(* CODESYS project keyence_sr.library
   Company: KOSTAL GmbH & Co.KG
   Version: 1.0.0.0
   DefaultNamespace: KOSTAL.AF2024.Drivers.Scanner.Keyence_SR
   Title: KOSTAL.AF2024.Drivers.Scanner.Keyence_SR
   Placeholder: KOSTAL.AF2024.Drivers.Scanner.Keyence_SR
   Author: Frank Dümpelmann
   DocFormat: reStructuredText

Project tree, tasks and I/O mapping:
  libraries: KOSTAL.AF2024.Core.ListOf, 1.0.0.0 (KOSTAL GmbH & Co.KG); KOSTAL.AF2024.Core.Process, 1.0.0.0 (KOSTAL GmbH & Co.KG); KOSTAL.AF2024.Core.Settings, 1.0.0.0 (KOSTAL GmbH & Co.KG); KOSTAL.AF2024.Core.StringTools, 1.0.0.0 (KOSTAL GmbH & Co.KG); KOSTAL.AF2024.Drivers.Scanner.IScanner, 1.0.0.0 (KOSTAL GmbH & Co.KG); Tc2_Standard, 3.3.3.0 (Beckhoff Automation GmbH); Tc2_TcpIp, 3.3.10.0 (Beckhoff Automation GmbH)
  DUT/
    data type E_PROCESS
  EthernetIP/
    DUTs/
      data type ST_SR751_IN
      data type ST_SR751_OUT
    function block FB_Reader_EthernetIP [ST]: ClearCodes, CodeGet, Ex_Scan, NativeStringGet, NumberOfBarcodes, State, _0_ready, _1_finish, _2_analyseResponse, _2_read, _2_split, _connectControl, _FBmain, FB_init, FBmain
  Project Information/
    function F_GetCompany [ST]
    function F_GetTitle [ST]
    function F_GetVersion [ST]
  TCP_IP/
    function block FB_Reader_TcpIp [ST]: ClearCodes, CodeGet, Ex_Scan, NativeStringGet, NumberOfBarcodes, State, _devices, _FBmain, _splitString, _stepConnect, _stepFinish, _stepReady, _stepReceive, _stepSend, _timeOutOccured, Command, ETX, ExecutedSocketState, intermediateLimiter, remote_IP, remote_Port, separator, serverAmsNetId, STX, timeOut, FB_init, FBmain
    interface I_Scanner: ExecutedSocketState
  Version/
    global variables Global_Version
*)

// DUT/E_PROCESS
{attribute 'qualified_only'}
{attribute 'strict'}
TYPE E_PROCESS :
(
	idle			:= 0,
	scan	:= 1
);
END_TYPE

// EthernetIP/DUTs/ST_SR751_IN
{attribute 'pack_mode' := '1'} 
TYPE ST_SR751_IN :
	STRUCT
		Error	: BIT;
		ResultDataAvailable	: BIT;
		ResultDataStrobe	: BIT;
		noName_0_0	: BIT;
		noName_0_1	: BIT;
		noName_0_2	: BIT;
		BufferOverfolwError	: BIT;
		GeneralError	: BIT;
		Busy	: BIT;
		TRG_BUSY	: BIT;
		LOCK_BUSY	: BIT;
		MODE_BUSY	: BIT;
		ERR_BUSY	: BIT;
		noName_1_0	: BIT;
		noName_1_1	: BIT;
		noName_1_2	: BIT;
		ReadComplete	: BIT;
		PresetComplete	: BIT;
		RegisterPresetDataComplete	: BIT;
		TuneComplete	: BIT;
		noName_2_0	: BIT;
		noName_2_1	: BIT;
		noName_2_2	: BIT;
		EXT_RequestComplete	: BIT;
		ReadFailure	: BIT;
		PresetFailure	: BIT;
		RegisterPresetDataFailure	: BIT;
		TuneFailure	: BIT;
		noName_3_0	: BIT;
		noName_3_1	: BIT;
		noName_3_2	: BIT;
		EXT_RequestFailure	: BIT;
		IN_1_Status	: BIT;
		IN_2_Status	: BIT;
		noName_4_0	: BIT;
		noName_4_1	: BIT;
		OUT_1_Status	: BIT;
		OUT_2_Status	: BIT;
		OUT_3_Status	: BIT;
		noName_5	: BIT;
		Unstable	: BIT;
		MatchingLevelUnstable	: BIT;
		ISO_IEC_15415_Unstable	: BIT;
		AIM_DPM_Unstable	: BIT;
		SAE_A59132_Unstable	: BIT;
		noName_6_0	: BIT;
		noName_6_1	: BIT;
		noName_6_2	: BIT;
		noName_6_3	: BIT;
		noName_6_4	: BIT;
		noName_6_5	: BIT;
		noName_6_6	: BIT;
		noName_6_7	: BIT;
		noName_6_8	: BIT;
		noName_6_9	: BIT;
		noName_6_10	: BIT;
		noName_6_11	: BIT;
		noName_6_12	: BIT;
		noName_6_13	: BIT;
		noName_6_14	: BIT;
		noName_6_15	: BIT;
		noName_6_16	: BIT;
		noName_6_17	: BIT;
		noName_6_18	: BIT;
		MatchingLevel	: UINT;
		ISO_IEC_15415_Grade	: UINT;
		AIM_DPM_Grade	: UINT;
		noName_7	: ARRAY[0..1] OF BYTE;
		ReadResultCode	: UINT;
		PresetResultCode	: UINT;
		RegisterPresetDataResultCode	: UINT;
		TuneResultCode	: UINT;
		noName_8	: ARRAY[0..5] OF BYTE;
		EXT_RequestResultCode	: UINT;
		GeneralErrorCode	: UINT;
		noName_9	: ARRAY[0..1] OF BYTE;
		ResultDataReadyCount	: UINT;
		ResultDataUpdateCount	: UINT;
		noName_10	: ARRAY[0..1] OF BYTE;
		ResultDataSize	: UINT;
		ResultData : STRING(81);
		
		
		
		
	END_STRUCT
END_TYPE

// EthernetIP/DUTs/ST_SR751_OUT

TYPE ST_SR751_OUT :
	STRUCT
		noName0_BIT	: BIT;
		ResultDataLatch	: BIT;
		noName_1_0	: BIT;
		noName_1_1	: BIT;
		noName_1_2	: BIT;
		noName_1_3	: BIT;
		noName_1_4	: BIT;
		ErrorClear	: BIT;
		ReadRequest	: BIT;
		PresetRequest	: BIT;
		RegisterPresetDataRequest	: BIT;
		TuneRequest	: BIT;
		noName_2_0	: BIT;
		noName_2_1	: BIT;
		noName_2_2	: BIT;
		noName_2_3	: BIT;
		ReadCompleteClear	: BIT;
		PresetCompleteClear	: BIT;
		RegisterPresetDataCompleteClear	: BIT;
		TuneCompleteClear	: BIT;
		noName_3_0	: BIT;
		noName_3_1	: BIT;
		noName_3_2	: BIT;
		ExtRequestCompleteClear	: BIT;
		noName_4	: BYTE;
		BankNumber	: UINT;
		noName_5_0	: BYTE;
		noName_5_1	: BYTE;
		noName_5_2	: BYTE;
		noName_5_3	: BYTE;
		UserDataSize:	UINT;
		UserData	: ARRAY[14..77] OF BYTE;
	END_STRUCT
END_TYPE

// Version/Global_Version
{attribute 'TcGenerated'}
{attribute 'no-analysis'}
{attribute 'linkalways'}
// This function has been automatically generated from the project information.
VAR_GLOBAL CONSTANT
	{attribute 'const_non_replaced'}
	stLibVersion_KOSTAL_AF2024_Drivers_Scanner_Keyence_SR : ST_LibVersion := (iMajor := 1, iMinor := 0, iBuild := 0, iRevision := 0, nFlags := 0, sVersion := '1.0.0.0');
END_VAR

// EthernetIP/FB_Reader_EthernetIP
(*
From EDS Specification Keyence_1003_0101.eds from 22.11.2012 12:56
===================================================================
*)

FUNCTION_BLOCK FB_Reader_EthernetIP IMPLEMENTS KOSTAL_AF2024_Drivers_Scanner_IScanner.I_Scanner



VAR
	ECatState	AT %I*	: UINT;	//link to EtherCat State from {Device x (ECAT EIP Scanner (EL6652))}.Inputs.State
	SR_750_Series_State	AT %I*	: UINT;	//link to {SR-750 Series}.Inputs.State

	SR751_IN	AT %I*	: ARRAY[2..173] OF BYTE; //link with Continious mode ATTENTION be sure, that the Array-Nodes are collapsed
	SR751_OUT	AT %Q*	: ARRAY[2..77] OF BYTE; //link with Continious mode ATTENTION be sure, that the Array-Nodes are collapsed
	
	_pIN		: POINTER TO ST_SR751_IN;
	_pOUT	: POINTER TO ST_SR751_OUT;

	//
	_step		: KOSTAL_AF2024_Core_Process.FB_processStep;
	_THIS_CALLED			: E_PROCESS;
	_THIS_IN_PROCESS		: E_PROCESS;
	_state 	: KOSTAL_AF2024_Core_Process.T_plcState;

	//
	_split	: Kostal_AF2024_Core_StringTools.FB_Split_UTF8;
	_barcodes	: KOSTAL_AF2024_Core_ListOf.FB_ListOfString_UTF8;
	
	_nativeResult	: KOSTAL_AF2024_Core_Settings.T_MaxString_UTF8;
	

	
END_VAR

VAR CONSTANT
	_DELIMITER	: STRING(1):= '$1D';
	_STX	: STRING(1):= '$02';
	_ETX	: STRING(1):= '$03';
	_CR	: STRING(1):= '$0D';
	_LF	: STRING(1):= '$0A';
END_VAR

METHOD ClearCodes

_barcodes.clear();
_nativeResult := '';
END_METHOD

METHOD CodeGet : STRING(255)
VAR_INPUT
	number	: UINT;
END_VAR
CodeGet:= _barcodes.line_GET(number);
END_METHOD

METHOD Ex_Scan : BOOL
IF _THIS_CALLED <> E_PROCESS.idle THEN //Another process is running: don't start this process!
	Ex_Scan:= FALSE;	
	RETURN; 
END_IF


_THIS_CALLED := E_PROCESS.scan;

_FBmain();	//Call sequence via _FBmain

Ex_Scan := _THIS_CALLED = _THIS_IN_PROCESS;	//Return true when process was started
END_METHOD

METHOD NativeStringGet : STRING(255)
NativeStringGet:= _nativeResult;
END_METHOD

PROPERTY PUBLIC NumberOfBarcodes : UDINT
GET
NumberOfBarcodes:= _barcodes.NumberOfLines;
END_GET
END_PROPERTY

PROPERTY State : KOSTAL_AF2024_Core_Process.I_T_plcState
GET

State := _state;
END_GET
END_PROPERTY

METHOD PROTECTED _0_ready
VAR_INPUT
END_VAR


IF _pOUT^.ReadRequest THEN _pOUT^.ReadRequest:= FALSE;	END_IF
_pOUT^.ReadCompleteClear:= _pIN^.ReadComplete OR _pIN^.ReadFailure;
 
_state.clear();

IF _pIN^.ReadComplete OR _pIN^.ReadFailure THEN
	_state.busy := TRUE;
	_state.description:= "wait until Scanner is not longer busy";
ELSE
	_step.INC();
END_IF
END_METHOD

METHOD PROTECTED _1_finish
VAR_INPUT
END_VAR

_state.clear();

_state.finish := TRUE;
_state.pass:= TRUE;

//IF NOT _startProcess THEN	_step.set(0);	END_IF
END_METHOD

METHOD PROTECTED _2_analyseResponse
VAR_INPUT
END_VAR

_pOUT^.ReadRequest:= FALSE;
 
_state.clear();
_state.busy := TRUE;

IF NOT _pIN^.ReadFailure THEN

	_step.INC();


ELSE
	
	
	_state.finish := TRUE;
	_state.fail:= TRUE;
	_state.description:= STRING_TO_WSTRING(_pIN^.ResultData);

END_IF
END_METHOD

METHOD PROTECTED _2_read
VAR_INPUT
END_VAR


_pOUT^.ReadRequest:= TRUE;
 
_state.clear();
_state.busy := TRUE;

IF NOT _pIN^.ReadComplete THEN

	_state.description:= "wait until Scanner is finish";
	
ELSE
	
	_nativeResult:= _pIN^.ResultData;
	_step.INC();
	
END_IF
END_METHOD

METHOD PROTECTED _2_split
VAR_INPUT
END_VAR

VAR
	_i: UDINT;
	_replace: STRING(255);
END_VAR


_split.clear();
_split.Delimiter:= _DELIMITER;
_split.split(_nativeResult);
_barcodes.clear();

FOR _i:= 1 TO _split.Results.NumberOfLines DO

	_replace:= _split.Results.line_GET(_i);

	IF _replace <> '' THEN
		_replace:= Kostal_AF2024_Core_StringTools.F_Replace_UTF8(source:= _replace,toReplace:= _STX, replaceWith:= '', numberOfReplaces:= -1);
		_replace:= Kostal_AF2024_Core_StringTools.F_Replace_UTF8(source:= _replace,toReplace:= _ETX, replaceWith:= '', numberOfReplaces:= -1);
		_replace:= Kostal_AF2024_Core_StringTools.F_Replace_UTF8(source:= _replace,toReplace:= _CR, replaceWith:= '', numberOfReplaces:= -1);
		_replace:= Kostal_AF2024_Core_StringTools.F_Replace_UTF8(source:= _replace,toReplace:= _LF, replaceWith:= '', numberOfReplaces:= -1);
		_barcodes.addLine(_replace);
		
	END_IF

END_FOR

_step.INC();
END_METHOD

METHOD PROTECTED _connectControl : BOOL
VAR_INPUT
END_VAR

 
IF ECatState <> 0  THEN

	_connectControl:= FALSE;

	_state.clear();
	_state.fail:= TRUE;
	_state.description:= Tc2_Standard.WCONCAT(UINT_TO_WSTRING(ECatState), ";Error from EtherCAT (EIP-Scanner)");


	_step.init();

ELSIF SR_750_Series_State <> 0 THEN

	_connectControl:= FALSE;

	_state.clear();
	_state.fail:= TRUE;
	_state.description:= Tc2_Standard.WCONCAT(UINT_TO_WSTRING(SR_750_Series_State), ";Error from Ethernet IP Connection");

	_step.init();

ELSE
	
	_connectControl:= TRUE;

END_IF
END_METHOD

METHOD PROTECTED _FBmain
VAR_INPUT
END_VAR

_pIN:= ADR(SR751_IN[2]);
_pOUT:= ADR(SR751_OUT[2]);


IF NOT _connectControl() THEN RETURN;	END_IF

IF _THIS_CALLED <> _THIS_IN_PROCESS THEN
	_step.init();
END_IF

_THIS_IN_PROCESS:= _THIS_CALLED;

IF _THIS_CALLED = E_PROCESS.scan THEN

	_step.Header();
	
	CASE _step.actual OF
		
		0:	_0_ready();
		1:	_2_read();
		2:	_2_analyseResponse();
		3:	_2_split();
		4:	_1_finish();
		
	ELSE
		
		_state.clear();
		_state.fail:= TRUE;
		_state.description:= Tc2_Standard.WCONCAT(INT_TO_WSTRING(_step.actual), ". Step does not exist");
		
	END_CASE

ELSE
	_state.clear();
	_state.ready := TRUE;
END_IF
END_METHOD

METHOD FB_init : BOOL
VAR_INPUT
	bInitRetains : BOOL; // if TRUE, the retain variables are initialized (warm start / cold start)
	bInCopyCode : BOOL;  // if TRUE, the instance afterwards gets moved into the copy code (online change)
END_VAR

_pIN:= ADR(SR751_IN[2]);
_pOUT:= ADR(SR751_OUT[2]);
END_METHOD

METHOD PUBLIC FBmain
VAR_INPUT
END_VAR
IF _THIS_CALLED = E_PROCESS.idle THEN
	_FBmain();
END_IF

_THIS_CALLED:= E_PROCESS.idle;
END_METHOD

END_FUNCTION_BLOCK

// TCP_IP/I_Scanner
INTERFACE I_Scanner EXTENDS KOSTAL_AF2024_Drivers_Scanner_IScanner.I_Scanner

(*
Description
===========
| State of the TCP/IP connection
*)
PROPERTY PUBLIC ExecutedSocketState : E_SocketConnectionState
GET
END_GET
END_PROPERTY

END_INTERFACE

// Project Information/F_GetCompany
// This function has been automatically generated from the project information.
{attribute 'signature_flag' := '1073741824'}
{attribute 'TcGenerated'}
{attribute 'no-analysis'}
FUNCTION F_GetCompany : WSTRING
VAR_INPUT
	
END_VAR

F_GetCompany := "KOSTAL GmbH & Co.KG";

END_FUNCTION

// Project Information/F_GetTitle
// This function has been automatically generated from the project information.
{attribute 'signature_flag' := '1073741824'}
{attribute 'TcGenerated'}
{attribute 'no-analysis'}
FUNCTION F_GetTitle : WSTRING
VAR_INPUT
	
END_VAR

F_GetTitle := "KOSTAL.AF2024.Drivers.Scanner.Keyence_SR";

END_FUNCTION

// Project Information/F_GetVersion
// This function has been automatically generated from the project information.
{attribute 'signature_flag' := '1073741824'}
{attribute 'TcGenerated'}
{attribute 'no-analysis'}
FUNCTION F_GetVersion : ST_LibVersion
VAR_INPUT
	
END_VAR

F_GetVersion.iMajor := 1;
F_GetVersion.iMinor := 0;
F_GetVersion.iBuild := 0;
F_GetVersion.iRevision := 0;
F_GetVersion.sVersion := '1.0.0.0';
F_GetVersion.nFlags := 0;

END_FUNCTION

// TCP_IP/FB_Reader_TcpIp
{info 'The Beckhoff Library >TF6310-TCP-IP.exe< is needed'}
(*

:Author: Frank Dümpelmann <f.duempelmann@kostal.com>, Martin Hundt <m.hundt@kostal.com>
:Date: 2019-01-07

Function
========
| Extension of FB_Reader to connect to a barcode reader via TCP/IP
| Tested with Keyence SR 750 

Usage notes
===============
| Asyncronous function block: FBmain() method must be called cyclicly
| The Beckhoff Library >TF6310-TCP-IP.exe< is needed
| 	_mode_SR750	:	BOOL;	// use this mode with KEYENCE SR 750, because the command Acknowlede is not possible to disable.

Methods and Properties
======================
| See bottom of this document for a detailed description of each method or property
| Methods starting with an underline(_) are internally used and can be ignored by the user

| Usage sample: ..\Device\Scanner\scannerBestPractice
| Usage Keyence Template ..\Device\Scanner\Keyence_SR\Keyence SR-750.ptc .. \Keyence SR-1000.ptc

*)
FUNCTION_BLOCK PUBLIC FB_Reader_TcpIp  IMPLEMENTS I_Scanner
VAR_INPUT
END_VAR
VAR_OUTPUT
END_VAR

VAR
	

	_step			: KOSTAL_AF2024_Core_Process.FB_processStep;	
	_THIS_CALLED			: E_PROCESS;
	_THIS_IN_PROCESS		: E_PROCESS;
	            	
	_state 			: KOSTAL_AF2024_Core_Process.T_plcState;
	            	
	_Command		: STRING;	//STRING to define in FB_init()
	_STX			: STRING;	//STRING to define in FB_init()
	_ETX			: STRING;	//STRING to define in FB_init()
	_timeOut		: TIME	;	//TIME to define in FB_init()
	
	_receivedString	: KOSTAL_AF2024_Core_Settings.T_MaxString_UTF8;
	_split			: Kostal_AF2024_Core_StringTools.FB_Split_UTF8;
	_barcodes		: KOSTAL_AF2024_Core_ListOf.FB_ListOfString_UTF8;

	_serverAmsNetId	: STRING:= '';	//STRING:= '' - default on local system
	_remote_IP			: STRING;	//STRING
	_remote_Port		: UDINT:= 9004;	//UDINT

	_socket				: Tc2_TcpIp.FB_ClientServerConnection;	//Tc2_TcpIp.FB_ClientServerConnection
	_executedSocketState	:	E_SocketConnectionState;
	
	_send			: Tc2_TcpIp.FB_SocketSend;	//Tc2_TcpIp.FB_SocketSend
	_receive	: Tc2_TcpIp.FB_SocketReceive;	//Tc2_TcpIp.FB_SocketReceive
	_receiveComponent	: STRING(255);	//STRING(255)
	_receiveAck	: STRING(255);	//STRING(255)

	_timeOutTimer	: TON;	//TON

	_intermediateLimiter	: STRING(1):= '$1D';
	_separator						: STRING(1):= '$1E';
	
	_subStep	: KOSTAL_AF2024_Core_Process.FB_processStep;
	_concat	: Kostal_AF2024_Core_StringTools.FB_Concat;
	
	
	

END_VAR

METHOD ClearCodes

_barcodes.clear();
_receivedString := '';
END_METHOD

(*
Description
===========
| get barcode element (number)
*)
METHOD CodeGet : KOSTAL_AF2024_Core_Settings.T_MaxString_UTF8
VAR_INPUT
	number	: UINT;
END_VAR
IF (number = 0) OR (number > _barcodes.numberOfLines) THEN
	CodeGet:= '';
ELSE
	CodeGet:= _barcodes.line_GET(number);
END_IF
END_METHOD

METHOD Ex_Scan : BOOL
IF _THIS_CALLED <> E_PROCESS.idle THEN //Another process is running: don't start this process!
	Ex_Scan:= FALSE;	
	RETURN; 
END_IF


_THIS_CALLED := E_PROCESS.scan;

_FBmain();	//Call sequence via _FBmain

Ex_Scan := _THIS_CALLED = _THIS_IN_PROCESS;	//Return true when process was started
END_METHOD

METHOD NativeStringGet : STRING(255)
NativeStringGet:= _receivedString;
END_METHOD

PROPERTY NumberOfBarcodes : UDINT
GET
NumberOfBarcodes:= _barcodes.NumberOfLines;
END_GET
END_PROPERTY

(*
Description
===========
| Status of the block
*)
PROPERTY PUBLIC State : KOSTAL_AF2024_Core_Process.I_T_plcState
GET


State := _state;
END_GET
END_PROPERTY

METHOD PROTECTED _devices
VAR_INPUT
END_VAR


_timeOutTimer(IN:= , PT:= _timeOut, Q=> , ET=> );

_socket
	(
		sSrvNetID	:= _serverAmsNetId, 
		nMode			:= Tc2_TcpIp.CONNECT_MODE_ENABLEDBG, 

		sRemoteHost	:= _remote_IP, 
		nRemotePort	:= _remote_Port, 

		bEnable			:= , 
		tReconnect	:= _timeOut, 

		bBusy		=> , 
		bError	=> , 
		nErrId	=> , 
		hSocket	=> , 
		eState	=> 
	);
	
IF _socket.bEnable THEN	_executedSocketState:= _socket.eState;	END_IF
	
_send
	(
		sSrvNetId	:= _serverAmsNetId, 
		hSocket		:= _socket.hSocket, 
		cbLen			:= INT_TO_UDINT(Tc2_Standard.LEN(_Command)), 
		pSrc			:= ADR(_Command), 
		bExecute	:= , 
		tTimeout	:= _timeOut, 

		bBusy			=> , 
		bError		=> , 
		nErrId		=> 
	);
	
	
	_receive
	(
		sSrvNetId	:= _serverAmsNetId, 
		hSocket		:= _socket.hSocket, 

		cbLen:= SIZEOF(_receiveComponent) - 1, 
		pDest:= ADR(_receiveComponent), 

		bExecute:= , 
		tTimeout:= _timeOut, 

		bBusy			=> , 
		bError		=> , 
		nErrId		=> , 
		nRecBytes	=> 
	);
END_METHOD

(*
Decription
==========
| To be called cyclicly, e.g. in DeviceDefine
*)
METHOD PROTECTED _FBmain
VAR_INPUT
END_VAR
IF _THIS_CALLED <> _THIS_IN_PROCESS THEN
	_step.init();
END_IF

_THIS_IN_PROCESS:= _THIS_CALLED;

IF _THIS_CALLED = E_PROCESS.scan THEN
	_step.Header();
	
	CASE _step.actual OF
	
		0:	_stepReady();
		1:	_stepConnect();
		2:	_stepSend();
		3:	_stepReceive();
		4:	_stepFinish();
	
	ELSE
		
		_state.clear();
		_state.description:= Tc2_Standard.WCONCAT("Step does not exist", INT_TO_WSTRING(_step.actual));
		_state.fail		:= TRUE;
		_state.finish	:= TRUE;
	
	END_CASE

ELSE
	_step.init();
	_state.clear();
	_state.ready := TRUE;
END_IF
_devices();
END_METHOD

(*
| split received string depends of STX ETX
*)
METHOD PROTECTED _splitString  : BOOL

VAR
	_i: UDINT;
	_element: STRING(255);
	_stxPos: INT;
	_code: STRING(255);
END_VAR


_barcodes.clear();

IF _receivedString = '' THEN
	
	;	// no splitting possible

	
// if EXT is defined
// ============================================================================
ELSIF _ETX <> '' THEN

	_split.clear();
	_split.Delimiter:= _ETX;
	_split.Split(_receivedString);

	// if additional STX is defined then select
	IF _STX <> '' THEN

		FOR _i:= 1 TO _split.Results.NumberOfLines DO
			
			_element:= _split.Results.line_GET(_i);
			_stxPos:= Tc2_Standard.FIND(STR1:= _element, STR2:= _STX);

			IF _stxPos > 0 THEN
				_barcodes.addLine(newLine:= Tc2_Standard.RIGHT(STR:= _element, SIZE:= Tc2_Standard.LEN( STR:= _element) - _stxPos ));
			END_IF
		END_FOR
	
	// no STX defined
	ELSE

		FOR _i:= 1 TO _split.Results.NumberOfLines DO
			_barcodes.addLine(_split.Results.line_GET(_i));
		END_FOR
	
	END_IF

	
// if only STX is defined
// ============================================================================
ELSIF _STX <> '' THEN
	
	_split.clear();
	_split.Delimiter:= _STX;
	_split.Split(_receivedString);

	FOR _i:= 1 TO _split.Results.NumberOfLines DO
		_barcodes.addLine(_split.Results.line_GET( _i));
	END_FOR

// neither STX or ETX is defined then no splitting possible
// ============================================================================
ELSE

	_barcodes.addLine(newLine:= _receivedString);

END_IF

_splitString:= _barcodes.NumberOfLines > 0;



IF _barcodes.NumberOfLines = 1 THEN

	_code:= _barcodes.line_GET(1);

	_split.clear();
	_split.Delimiter:= _intermediateLimiter;
	_split.split(_code);

	_barcodes.removeLine(1);

	FOR _i:= 1 TO _split.Results.NumberOfLines DO
		_barcodes.addLine(_split.Results.line_GET(_i));
	END_FOR


END_IF
END_METHOD

METHOD PROTECTED _stepConnect
VAR_INPUT
END_VAR

IF _step.toggle THEN
	_state.clear();
	_state.busy:= TRUE;
	_subStep.init();
END_IF


IF _timeOutTimer.Q THEN

	_timeOutOccured();

ELSE

	_subStep.Header();
	
	CASE _subStep.actual OF
		0:	_socket.bEnable:= FALSE;	_subStep.INC();
		1:	_socket.bEnable:= TRUE;		_subStep.INC();

		2:	IF _socket.bBusy THEN
					_state.busy	:= TRUE;
					_state.description:= "Scanner is busy(connect); wait ...";
				ELSE
					_subStep.INC();
				END_IF

		3:	IF _socket.bError THEN
					_state.clear();
					_state.description:= Tc2_Standard.WCONCAT("Error during socket open. Errorcode>", UDINT_TO_WSTRING(_socket.nErrId));
					_state.fail	:= TRUE;
					_state.finish:= TRUE;	
					_timeOutTimer.IN:= FALSE;
				ELSIF _socket.hSocket.handle = 0 THEN
					_state.clear();
					_state.description:= "no Handle from socket";
					_state.fail	:= TRUE;
					_state.finish:= TRUE;
					_timeOutTimer.IN:= FALSE;
				ELSE
					_step.INC();
				END_IF
		
	ELSE
	
		_timeOutTimer.IN:= FALSE;
		_state.clear();
		_state.fail	:= TRUE;
		_state.finish:= TRUE;
		_concat.clear();
		_concat.addContent("connect Step ");
		_concat.addContent(INT_TO_WSTRING(_subStep.actual));
		_concat.addContent(" does not exist");
		_state.description:= _concat.getResult();
		_concat.clear();
	
	END_CASE

END_IF
END_METHOD

METHOD PROTECTED _stepFinish
VAR_INPUT
END_VAR

IF _step.toggle THEN

	_timeOutTimer.IN:= FALSE;

	_socket.bEnable		:= FALSE;
	_send.bExecute		:= FALSE;
	_receive.bExecute	:= FALSE;

END_IF

_state.busy		:= FALSE;
_state.finish	:= TRUE;
END_METHOD

METHOD PROTECTED _stepReady
VAR_INPUT
END_VAR

IF _step.toggle THEN

	_state.clear();
	_state.ready		:= TRUE;

	_socket.bEnable		:= FALSE;
	_send.bExecute		:= FALSE;
	_receive.bExecute	:= FALSE;

	_timeOutTimer.IN:= FALSE;

END_IF


IF NOT _step.toggle THEN

	_step.INC();

	_receivedString:= '';
	_receiveComponent:= '';
	
	_receiveAck:= '';

	_split.clear();
	_barcodes.clear();
	
	_timeOutTimer.IN:= TRUE;
	
	_state.clear();
	_state.busy:= TRUE;

ELSE

	_state.clear();
	_state.ready:= TRUE;
		
END_IF
END_METHOD

METHOD PROTECTED _stepReceive
VAR_INPUT
END_VAR

IF _step.toggle THEN

	_state.clear();
	_state.busy:= TRUE;

	_subStep.init();

	_receivedString:= '';
	_receiveComponent:= '';

	_split.clear();
	_barcodes.clear();

END_IF



IF _timeOutTimer.Q THEN

	_timeOutOccured();

ELSE
	
	_subStep.Header();

	CASE _subStep.actual OF
		0:	_receive.bExecute:= FALSE;	_receiveComponent:= '';	_subStep.INC();
		1:	_receive.bExecute:= TRUE;		_subStep.INC();

		2:	IF _receive.bBusy THEN
					_state.busy	:= TRUE;
					_state.description:= "Scanner is busy(receive); wait ...";
				ELSE
					_subStep.INC();
				END_IF

		3:	IF _receive.bError THEN
					_state.clear();
					_state.description:= Tc2_Standard.WCONCAT("Error during receive. Errorcode>", UDINT_TO_WSTRING(_receive.nErrId));
					_state.fail	:= TRUE;
					_state.finish:= TRUE;	
					_timeOutTimer.IN:= FALSE;
				ELSE
					_subStep.INC();
				END_IF
		
		4:	IF	_receive.nRecBytes <> 0 THEN 

					_receivedString:= Tc2_Standard.CONCAT(STR1:= _receivedString, STR2:=  Tc2_Standard.LEFT(STR:= _receiveComponent, SIZE:= UDINT_TO_INT(_receive.nRecBytes)));
					_receiveComponent:= '';
					_splitString();

					_subStep.SET(0);

				ELSIF _barcodes.NumberOfLines < 1 THEN 

					_subStep.SET(0);

				ELSE
					
					_state.clear();
					_state.busy:= TRUE;
					_state.pass:= TRUE;
					_timeOutTimer.IN:= FALSE;
					_step.INC();

				END_IF
								
	ELSE
	
		_timeOutTimer.IN:= FALSE;
		_state.clear();
		_state.fail	:= TRUE;
		_state.finish:= TRUE;
		_concat.clear();
		_concat.addContent("send Step ");
		_concat.addContent(INT_TO_WSTRING(_subStep.actual));
		_concat.addContent(" does not exist");
		_state.description:= _concat.getResult();
		_concat.clear();
	
	END_CASE

END_IF
END_METHOD

METHOD PROTECTED _stepSend
VAR_INPUT
END_VAR

IF _step.toggle THEN
	_state.clear();
	_state.busy:= TRUE;
	_subStep.init();
END_IF


IF _timeOutTimer.Q THEN

	_timeOutOccured();

ELSE
	
	_subStep.Header();

	CASE _subStep.actual OF
		0:	_send.bExecute:= FALSE;	_subStep.INC();
		1:	_send.bExecute:= TRUE;		_subStep.INC();

		2:	IF _send.bBusy THEN
					_state.busy	:= TRUE;
					_state.description:= "Scanner is busy(send); wait ...";
				ELSE
					_subStep.INC();
				END_IF

		3:	IF _send.bError THEN
					_state.clear();
					_state.description:= Tc2_Standard.WCONCAT("Error during send. Errorcode>", UDINT_TO_WSTRING(_send.nErrId));
					_state.fail	:= TRUE;
					_state.finish:= TRUE;	
					_timeOutTimer.IN:= FALSE;
				ELSE
					_step.INC();
				END_IF
		
	ELSE
	
		_state.clear();
		_state.fail	:= TRUE;
		_state.finish:= TRUE;
		_concat.clear();
		_concat.addContent("send Step ");
		_concat.addContent(INT_TO_WSTRING(_subStep.actual));
		_concat.addContent(" does not exist");
		_state.description:= _concat.getResult();
		_concat.clear();
	
	END_CASE

END_IF
END_METHOD

METHOD PROTECTED _timeOutOccured
VAR_INPUT
END_VAR


_socket.bEnable		:= FALSE;
_send.bExecute		:= FALSE;
_receive.bExecute	:= FALSE;

_state.busy:= FALSE;
_state.description:= "Timeout";
_state.fail:= TRUE;
_state.finish:= TRUE;
END_METHOD

(*
Description
===========
| Command to start scanner
| default: t$0D$0A
*)
PROPERTY PUBLIC Command : String
GET

Command:= _Command;
END_GET
SET

_Command:= Command;
END_SET
END_PROPERTY

(*
Description
===========
| 'End of text' command in the string from the reader
| default: $03
*)
PROPERTY PUBLIC ETX : String
GET

ETX:= _ETX;
END_GET
SET

_ETX:= ETX;
END_SET
END_PROPERTY

(*
Description
===========
| State of the TCP/IP connection
*)
PROPERTY PUBLIC ExecutedSocketState : E_SocketConnectionState
GET

ExecutedSocketState:= _executedSocketState;
END_GET
END_PROPERTY

PROPERTY PUBLIC intermediateLimiter : STRING(1)
GET

intermediateLimiter:= _intermediateLimiter;
END_GET
SET

_intermediateLimiter:= intermediateLimiter;
END_SET
END_PROPERTY

(*
Description
===========
| IP address of the barcode reader
*)
PROPERTY PUBLIC remote_IP : STRING
GET


remote_IP:= _remote_IP;
END_GET
SET

_remote_IP:= remote_IP;
END_SET
END_PROPERTY

(*
Description
===========
| TCP/IP port of the barcode reader
*)
PROPERTY PUBLIC remote_Port : UDINT
GET


remote_Port:= _remote_Port;
END_GET
SET

_remote_Port:= remote_Port;
END_SET
END_PROPERTY

PROPERTY PUBLIC separator : STRING(1)
GET

separator:= _separator;
END_GET
SET

_separator:= separator;
END_SET
END_PROPERTY

(*
Description
===========
| AmsNetId of the system running the Beckhoff TCP/IP server
| default: ''=local system
*)
PROPERTY PUBLIC serverAmsNetId : STRING
GET

serverAmsNetId:= _serverAmsNetId;
END_GET
SET

_serverAmsNetId:= serverAmsNetId;
END_SET
END_PROPERTY

(*
Description
===========
| 'Start of text' command in the string from the reader
| default: $02
*)
PROPERTY PUBLIC STX : String
GET

STX:= _STX;
END_GET
SET

_STX:= STX;
END_SET
END_PROPERTY

(*
Description
===========
| Time after fault is generated when scanner does not respond
| default: 5s
*)
PROPERTY PUBLIC timeOut : TIME
GET

timeOut:= _timeOut;
END_GET
SET

IF timeOut > T#0MS THEN
	_timeOut:= timeOut;
END_IF
END_SET
END_PROPERTY

METHOD FB_init : BOOL
VAR_INPUT
	bInitRetains : BOOL; // if TRUE, the retain variables are initialized (warm start / cold start)
	bInCopyCode : BOOL;  // if TRUE, the instance afterwards gets moved into the copy code (online change)
END_VAR

_Command	:= 'LON$0D';	//STRING	:= 'LON$R'
_STX			:= '$02';			//STRING	:= '$02'
_ETX			:= '$03';			//STRING	:= '$03'
_timeOut	:= T#5S;			//TIME:= T#5S - default

_intermediateLimiter:= '$1D';
_separator					:= '$1E';
END_METHOD

METHOD PUBLIC FBmain
VAR_INPUT
END_VAR
IF _THIS_CALLED = E_PROCESS.idle THEN
	_FBmain();
END_IF

_THIS_CALLED:= E_PROCESS.idle;
END_METHOD

END_FUNCTION_BLOCK
